(*
SPDX-FileCopyrightText: © 2026 Oleksandr Tiutyk <trofimich@gmail.com>
SPDX-License-Identifier: MIT
License: https://opensource.org/license/mit
*)

(*!
<summary>Holds a multi-field live value for native JSON round-trip tests.</summary>
*)
TYPE JSON_TEST_VALUE :
STRUCT
	//! <summary>Integer payload with an independent expected value.</summary>
	Number : DINT;
	//! <summary>Boolean payload used to detect incomplete restoration.</summary>
	Ready : BOOL;
END_STRUCT
END_TYPE

(* stored: Version 1.1.0.1
   DUT JSON_TEST_VALUE: Id {7289aec6-4f4e-4ecc-a209-5b1b102147d1} *)
